Fanuc KAREL source: ko00036.KL

-- PROVISIONAL review KL for V770-1; original PC SHA256 8ad17e90a4f891a48a5a20a3c3379bdc1c53a56efd56d2f109707be1a8c372ad
-- Incomplete behavior may be omitted. Consult companion uncertainty JSON. Do not deploy.
PROGRAM KO00036
%NOLOCKGROUP
BEGIN
  -- UNRESOLVED_PC offsets 5-12; opcodes 9D,23
  -- UNRESOLVED_PC offsets 17-66; opcodes 27,27,49,7E,AD,22,1C,22,31,7E,4A
  -- UNRESOLVED_PC offsets 71-75; opcodes 7F
END KO00036
